(* PLC project Vn_move_stmt, Beckhoff Automation GmbH TwinCAT PLC Control 3.5.13.21 *)
(* stored: creationDateTime 1970-01-01T00:00:00 *)

PROGRAM Vn_move_stmt

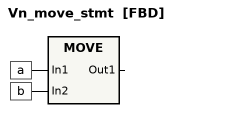
(* FBD diagram, written out as Structured Text *)
MOVE(a, b);
END_PROGRAM
